SUBAPPLICATION FU_Demo_H300 (* Ein DELIXI H300 (0,75 kW) per Modbus RTU hinter einem Waveshare RS232/485/422 TO POE ETH (B) (Modbus TCP<->RTU, Port 502). Messwerte: der Modbus-Client pollt selbst alle 500 ms und meldet jede Abfrage per CNF; skalieren, auf den lokalen OPC-UA-Server publizieren. Kommando: Steuerwort vom Web-Dashboard -> 9300H (genau ein Write je Dashboard-Klick). Sollwert: Sollfrequenz in Hz vom Web-Dashboard -> begrenzen -> % von Fmax -> 9301H. Nur Standard-/logiBUS-Typen, die auf der APIXON bereits als ELF-Lib vorhanden sind - kein eigener FB-Typ, kein Firmware-Build noetig. *)
  (* Standard: 61499-2; Description: Copyright (c) 2026 Franz Höpfinger This program and the accompanying materials are made available under the terms of the Eclipse Public License 2.0 which is available at https://www.eclipse.org/legal/epl-2.0/ SPDX-License-Identifier: EPL-2.0 *)
  (* Version 1.2, 2026-11-02, Franz Höpfinger, Franz Höpfinger, Ticker (MyLib::sys::SystemTickSender_OPC): Lebenszeichen FU1.SYSTEM_TICK fuer das Dashboard. *)
  (* Version 1.1, 2026-11-02, Franz Höpfinger, Franz Höpfinger, in drei SubApps aufgeteilt (FU_Messwerte, FU_Kommando, FU_Sollwert), E_CYCLE entfernt *)
  (* Version 1.0, 2026-11-02, Franz Höpfinger, Franz Höpfinger, initial *)
  PACKAGE FBs::FU_Demo;
  IMPORT FBs::FU_Demo::FU_Demo_Konstanten::FU_SYSTEM_TICK_WEB_WRITE;
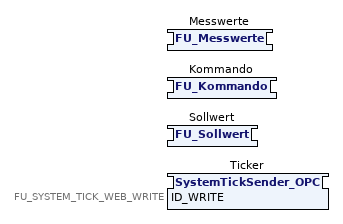
  SUBAPPS
    Messwerte : FBs::FU_Demo::FU_Messwerte;
    Kommando : FBs::FU_Demo::FU_Kommando;
    Sollwert : FBs::FU_Demo::FU_Sollwert;
    Ticker : MyLib::sys::SystemTickSender_OPC(ID_WRITE := FU_SYSTEM_TICK_WEB_WRITE); (* Lebenszeichen fuer das Web-Dashboard *)
  END_SUBAPPS
END_SUBAPPLICATION
